Yaskawa INFORM job: -DEFRO-70-PRZYLACZE-70-KOPIA-.JBI

/JOB
//NAME -DEFRO-70-PRZYLACZE-70-KOPIA-
//POS
///NPOS 40,40,40,0,0,0
///TOOL 0
///POSTYPE PULSE
///PULSE
C00000=-281,-101163,-84214,3730,-80188,-1936
C00001=-283,-101162,-84213,3710,-80188,-1936
C00002=116617,-39062,-41553,1138,-40446,20
C00003=97332,10008,-65831,-77395,-56626,78097
C00004=97332,10036,-65835,-77406,-56622,78106
C00005=126597,-12792,-74683,9116,-14112,37031
C00006=129578,-9389,-72169,26197,-17561,29790
C00007=143171,23000,-49885,51799,-48783,19450
C00008=142289,27625,-43624,46606,-52109,19593
C00009=140707,34961,-33804,39360,-57405,19440
C00010=137188,46732,-18219,29241,-65914,18506
C00011=125601,64166,5444,7463,-78162,8461
C00012=120628,60223,2537,-370,-74792,3762
C00013=116260,63341,4618,-6746,-77452,-573
C00014=112604,59060,-1014,-13680,-74421,-638
C00015=105645,46181,-18056,-25918,-65595,-11662
C00016=96917,44348,-31091,-45677,-66308,-16214
C00017=100527,41964,-28031,-34606,-66372,-26006
C00018=106433,45775,-18486,-19914,-75527,-46558
C00019=110224,24520,-34980,-16270,-62186,-56055
C00020=117116,19907,-37131,-3644,-59039,-60958
C00021=117137,19542,-37273,-3641,-59137,-60967
C00022=117062,4461,-25894,-3265,-73866,-61376
C00023=125074,-50101,-76658,51202,-17672,58606
C00024=125043,-41373,-84041,81327,-13668,44712
C00025=124776,-28424,-75745,87893,-13306,41755
C00026=124712,-28431,-75750,87904,-13268,41762
C00027=120787,-27884,-69765,25728,-8700,23794
C00028=115036,-25344,-64782,-26451,-15542,29683
C00029=119186,-28374,-69103,18427,-8940,-7851
C00030=122010,-28108,-68825,46224,-14319,-44839
C00031=116778,-25971,-65828,-246,-14948,-40490
C00032=118192,-23314,-61354,4708,-22161,-64875
C00033=115451,-27710,-69473,-21973,-12695,-70389
C00034=115429,-28374,-69925,-21919,-12759,-70410
C00035=115209,-37948,-70943,-16962,-16869,-72656
C00036=119279,-50675,-71302,9013,-26968,83196
C00037=116617,-39062,-41553,1138,-40446,20
C00038=-283,-101162,-84213,3710,-80188,-1936
C00039=-281,-101163,-84214,3730,-80188,-1936
BC00000=570125
BC00001=954451
BC00002=878037
BC00003=878036
BC00004=878036
BC00005=878037
BC00006=878037
BC00007=878037
BC00008=878037
BC00009=878037
BC00010=878037
BC00011=878037
BC00012=878036
BC00013=878037
BC00014=878037
BC00015=878037
BC00016=878037
BC00017=878037
BC00018=878037
BC00019=878037
BC00020=878037
BC00021=878037
BC00022=878037
BC00023=869720
BC00024=869720
BC00025=869720
BC00026=869720
BC00027=869721
BC00028=869721
BC00029=869721
BC00030=869721
BC00031=869721
BC00032=869721
BC00033=869721
BC00034=869721
BC00035=869721
BC00036=869720
BC00037=878037
BC00038=954451
BC00039=570125
EC00000=1163,0
EC00001=1166,0
EC00002=-1743,0
EC00003=-1746,0
EC00004=-1746,0
EC00005=-1743,0
EC00006=-1743,0
EC00007=-1743,0
EC00008=-1743,0
EC00009=-1743,0
EC00010=-1744,0
EC00011=-1744,0
EC00012=-1745,0
EC00013=-1744,0
EC00014=-1744,0
EC00015=-1744,0
EC00016=-1744,0
EC00017=-1744,0
EC00018=-1744,0
EC00019=-1744,0
EC00020=-1744,0
EC00021=-1744,0
EC00022=-1744,0
EC00023=-85617,0
EC00024=-85617,0
EC00025=-85617,0
EC00026=-85617,0
EC00027=-85617,0
EC00028=-85617,0
EC00029=-85617,0
EC00030=-85617,0
EC00031=-85617,0
EC00032=-85617,0
EC00033=-85617,0
EC00034=-85617,0
EC00035=-85617,0
EC00036=-85617,0
EC00037=-1743,0
EC00038=1166,0
EC00039=1163,0
//INST
///DATE 2026/09/14 21:41
///ATTR SC,RW
///GROUP1 RB1,BS1
///GROUP2 ST1
NOP
MOVJ C00000 BC00000 VJ=80.00 DEC=20  +MOVJ EC00000 VJ=80.00
MOVJ C00001 BC00001 VJ=80.00 DEC=20  +MOVJ EC00001 VJ=0.78
MOVJ C00002 BC00002 VJ=80.00 DEC=20  +MOVJ EC00002 VJ=80.00
MOVJ C00003 BC00003 VJ=80.00 DEC=20  +MOVJ EC00003 VJ=2.00
TIMER T=0.50
MACRO1 MJ#(0) ARGF8
ARCON
WVON WEV#(21)
MOVC C00004 BC00004 V=5.0 DEC=20  +MOVJ EC00004 VJ=80.00
MOVC C00005 BC00005 V=5.0 DEC=20  +MOVJ EC00005 VJ=80.00
MOVC C00006 BC00006 V=5.0 DEC=20  +MOVJ EC00006 VJ=80.00
MOVL C00007 BC00007 V=5.0 DEC=20  +MOVJ EC00007 VJ=80.00
MOVL C00008 BC00008 V=7.5 DEC=20  +MOVJ EC00008 VJ=80.00
MOVL C00009 BC00009 V=5.0 DEC=20  +MOVJ EC00009 VJ=0.78
MOVC C00010 BC00010 V=5.0 DEC=20  +MOVJ EC00010 VJ=80.00
MOVC C00011 BC00011 V=5.0 DEC=20  +MOVJ EC00011 VJ=80.00
WVON WEV#(22)
MOVC C00012 BC00012 V=5.0 DEC=20  +MOVJ EC00012 VJ=80.00
MOVC C00013 BC00013 V=5.0 DEC=20  +MOVJ EC00013 VJ=80.00
WVON WEV#(23)
MOVC C00014 BC00014 V=5.0 DEC=20  +MOVJ EC00014 VJ=80.00
MOVC C00015 BC00015 V=5.0 DEC=20  +MOVJ EC00015 VJ=80.00
MOVL C00016 BC00016 V=5.0 DEC=20  +MOVJ EC00016 VJ=80.00
MOVL C00017 BC00017 V=7.5 DEC=20  +MOVJ EC00017 VJ=80.00
WVON WEV#(21)
MOVC C00018 BC00018 V=6.7 DEC=20  +MOVJ EC00018 VJ=80.00
MOVL C00019 BC00019 V=5.0 DEC=20  +MOVJ EC00019 VJ=80.00
MOVL C00020 BC00020 V=5.0 DEC=20  +MOVJ EC00020 VJ=80.00
MOVC C00021 BC00021 V=5.0 DEC=20  +MOVJ EC00021 VJ=80.00
ARCOF
WVOF
MOVJ C00022 BC00022 VJ=80.00 DEC=20  +MOVJ EC00022 VJ=80.00
MOVJ C00023 BC00023 VJ=80.00 DEC=20  +MOVJ EC00023 VJ=80.00
MOVJ C00024 BC00024 VJ=80.00 DEC=20  +MOVJ EC00024 VJ=80.00
MOVJ C00025 BC00025 VJ=80.00 DEC=20  +MOVJ EC00025 VJ=80.00
TIMER T=0.50
MACRO1 MJ#(0) ARGF4
ARCON
MOVC C00026 BC00026 V=5.0 DEC=20  +MOVJ EC00026 VJ=80.00
MOVC C00027 BC00027 V=5.0 DEC=20  +MOVJ EC00027 VJ=80.00
MOVC C00028 BC00028 V=5.0 DEC=20  +MOVJ EC00028 VJ=80.00
MOVC C00029 BC00029 V=5.0 DEC=20  +MOVJ EC00029 VJ=80.00
MOVC C00030 BC00030 V=5.0 DEC=20  +MOVJ EC00030 VJ=80.00
MOVC C00031 BC00031 V=5.0 DEC=20  +MOVJ EC00031 VJ=80.00
MOVC C00032 BC00032 V=5.0 DEC=20  +MOVJ EC00032 VJ=80.00
MOVC C00033 BC00033 V=5.0 DEC=20  +MOVJ EC00033 VJ=80.00
MOVJ C00034 BC00034 VJ=2.00 DEC=20  +MOVJ EC00034 VJ=80.00
ARCOF
MOVJ C00035 BC00035 VJ=80.00 DEC=20  +MOVJ EC00035 VJ=80.00
MOVJ C00036 BC00036 VJ=80.00 DEC=20  +MOVJ EC00036 VJ=80.00
MOVJ C00037 BC00037 VJ=80.00 DEC=20  +MOVJ EC00037 VJ=80.00
MOVJ C00038 BC00038 VJ=80.00 DEC=20  +MOVJ EC00038 VJ=80.00
MOVJ C00039 BC00039 VJ=80.00 DEC=20  +MOVJ EC00039 VJ=80.00
END
